// TIA Portal V20 export
TYPE "Drehteller"
   STRUCT
      Wartungsintervall : DInt;
      Fertigmeldung_Drehteller : Bool;
      Aktorzyklen : DInt;
      Auto_Frg_Drehen_Vorwärts : Bool;
      Auto_Frg_Drehen_Rückwärts : Bool;
      Manu_Frg_Drehen_Vorwärts : Bool;
      Manu_Frg_Drehen_Rückwärts : Bool;
      Richt_Frg_Drehen_Vorwärts : Bool;
      Richt_Frg_Drehen_Rückwärts : Bool;
   END_STRUCT;
END_TYPE
